// TIA Portal V19 export
// export: Created 2026-10-15T10:10:34.3952238Z, ExportSetting WithDefaults, DisplayName Totally Integrated Automation Portal, DisplayVersion V19, DisplayName TIA Portal Openness, DisplayVersion V19, DisplayName TIA Portal Version Control Interface, DisplayVersion V19, DisplayName STEP 7 Professional, DisplayVersion V19, DisplayName STEP 7 Safety, DisplayVersion V19, DisplayName WinCC Basic/Comfort/Advanced, DisplayVersion V19, DisplayName WinCC Unified, DisplayVersion V19
DATA_BLOCK "ROLL_IO"   // DB2
{ S7_Optimized_Access := 'TRUE' }
VERSION : 0.1
// stored: AutoNumber true, DBAccessibleFromOPCUA true, DBAccessibleFromWebserver true, IsOnlyStoredInLoadMemory false, IsRetainMemResEnabled false, IsWriteProtectedInAS false, MemoryReserve 100
   VAR
      Input : Array[0..127, 0..7] of Bool;
      Output : Array[0..127, 0..7] of Bool;
      Simulation : Bool := TRUE;
      PhysicalOutputsEnabled : Bool := FALSE;
      PhysicalIoConfigured : Bool := FALSE;
      ConversionFault : Bool;
      FirstCycle : Bool := TRUE;
      RuntimeMemory : LReal;
      ClockMs : LReal;
      HmiElapsedMs : LReal;
      HmiLastHeartbeat : DInt;
   END_VAR
BEGIN
END_DATA_BLOCK
